Fanuc KAREL source: kx00029.KL

-- PROVISIONAL review KL for V770-1; original PC SHA256 712b45c482f98f27cde57f02bf66fb97911500fce2b850f887dc5ea4ad734ae7
-- Incomplete behavior may be omitted. Consult companion uncertainty JSON. Do not deploy.
PROGRAM KX00029
%NOLOCKGROUP
VAR
  I : INTEGER
  J : INTEGER
  B : BOOLEAN
  F : FILE
  S : STRING[80]
-- UNRESOLVED_DECL P type=000102
BEGIN
  -- UNRESOLVED_PC offsets 5-12; opcodes 9D,23
  -- UNRESOLVED_PC offsets 17-21; opcodes 7F
END KX00029
